(* IEC 61131-3 sources: veristc/veri-stc/tests/compiler-tests/positive, 6 files *)

(* ---- algo_blocks_fb.st ---- *)
(* ================================================================
   algo_blocks_fb.st
   原生 FUNCTION_BLOCK 版算法块库 + "不同变量调用相同算法功能" e2e

   与 FUNCTION 版（algo_blocks_lib.st / algo_blocks_multi_instance.st）
   同激励、同黄金时间线，可交叉验证两种实现一致。

   演示 FB 全部可用特性（P1 + v1.5）：
     - VAR_INPUT / VAR_OUTPUT（多输出：Q 与 QN、U 与 UI 与 ALM）
     - VAR 实例内持久状态（UI / E_OLD，FB_DATA 跨周期不清零）
     - VAR_IN_OUT 逐引用别名（TRACE：诊断量直写调用方全局）
     - 实例声明分离：rs1/rs2 同一份代码、独立数据段
     - IF/ELSIF/ELSE 控制流、表达式实参、命名实参（:=）
   限制：FB 体内不得声明成员实例（嵌套 FB 不支持，P1 范围外）。
   调用点在外部以 IEC 点号访问 inst.FIELD 读取字段（v1.5.1；编译器内部
   融合为不可书写的派生名 inst#FIELD，外部只能读 VAR_OUTPUT）。

   黄金时间线（数值列与 FUNCTION 版一致，t: rs1 rs2 sr1 sr2 | u1 ui1 |
   u2 ui2 | f1 f2，u 与 tr 恒等因 TRACE 别名）。列标签自 v1.5.1 起写作
   点号形式（rs1.Q / pid1.U / pid1.UI / fby1.Y …）指认"这一列来自哪个
   实例的哪个字段"；golden 文件随之只改标签文本，12 行数值逐列不变：
     t1 : 1 0 0 0 | 170 118 | 140 65  |  20   0
     t2 : 1 0 0 0 | 170 200 | 140 90  |  40   0
     t3 : 1 1 0 0 | 170 200 | 140 90  |  60   0
     t4 : 1 0 0 0 | 170 200 | 140 90  |  80   0
     t5 : 0 0 0 0 | 170 200 | 140 90  | 100  50
     t6 : 0 0 0 1 | 170 200 | 140 90  | 120 100
     t7 : 0 0 0 1 | 170 200 | 140 90  | 140 120
     t8 : 0 0 0 1 | 170 200 | 140 90  | 160 120
     t9 : 0 0 0 0 | 170 200 | 135 90  | 180 120
     t10: 0 0 0 0 | 170 200 | 125 90  | 200 120
     t11: 0 0 0 0 | 170 198 | 115 90  | 220 120
     t12: 0 0 0 0 | 158 184 | 105 90  | 240 120
   ================================================================ *)

(* ---- 实例声明：必须先于 POU 列表；每实例独立 FB_DATA ---- *)
VAR_GLOBAL
  rs1  : RS_FB;
  rs2  : RS_FB;
  sr1  : SR_FB;
  sr2  : SR_FB;
  pid1 : PID_FB;
  pid2 : PID_FB;
  fby1 : FBY_FB;
  fby2 : FBY_FB;
  trace1 : DINT;   (* pid1 的 VAR_IN_OUT 别名目标 *)
  trace2 : DINT;   (* pid2 的 VAR_IN_OUT 别名目标 *)
END_VAR

(* ---- RS：置位优先双稳态；Q 为实例持久状态 ---- *)
FUNCTION_BLOCK RS_FB
VAR_INPUT
  S : BOOL;
  R : BOOL;
END_VAR
VAR_OUTPUT
  Q  : BOOL;
  QN : BOOL;
END_VAR
  Q := S OR (Q AND NOT R);
  QN := NOT Q;
END_FUNCTION_BLOCK

(* ---- SR：复位优先双稳态 ---- *)
FUNCTION_BLOCK SR_FB
VAR_INPUT
  S : BOOL;
  R : BOOL;
END_VAR
VAR_OUTPUT
  Q  : BOOL;
  QN : BOOL;
END_VAR
  Q := (S OR Q) AND NOT R;
  QN := NOT Q;
END_FUNCTION_BLOCK

(* ---- PID：定点 PID，实例内持久 UI/E_OLD，KI 固定为 1；
       TRACE 为 VAR_IN_OUT 诊断别名，输出 U 同步写入调用方全局 ---- *)
FUNCTION_BLOCK PID_FB
VAR_INPUT
  E     : DINT;
  KP    : DINT;
  KD    : DINT;
  UI_LO : DINT;
  UI_HI : DINT;
  LO    : DINT;
  HI    : DINT;
END_VAR
VAR_OUTPUT
  U   : DINT;
  UI  : DINT;
  ALM : BOOL;
END_VAR
VAR_IN_OUT
  TRACE : DINT;
END_VAR
VAR
  DE    : DINT;
  V     : DINT;
  E_OLD : DINT;
END_VAR
  DE := E - E_OLD;
  V := UI + E;
  IF V > UI_HI THEN
    V := UI_HI;
  ELSIF V < UI_LO THEN
    V := UI_LO;
  END_IF;
  UI := V;
  U := KP * E + UI + KD * DE;
  IF U > HI THEN
    U := HI;
  ELSIF U < LO THEN
    U := LO;
  END_IF;
  IF U >= HI THEN
    ALM := TRUE;
  ELSE
    ALM := FALSE;
  END_IF;
  TRACE := U;
  E_OLD := E;
END_FUNCTION_BLOCK

(* ---- FBY：速率限制跟随；Y 为实例持久输出 ---- *)
FUNCTION_BLOCK FBY_FB
VAR_INPUT
  IN : DINT;
  DR : DINT;
END_VAR
VAR_OUTPUT
  Y : DINT;
END_VAR
VAR
  V : DINT;
END_VAR
  V := IN;
  IF V > Y + DR THEN
    V := Y + DR;
  ELSIF V < Y - DR THEN
    V := Y - DR;
  END_IF;
  Y := V;
END_FUNCTION_BLOCK

PROGRAM MAIN
VAR
  tick : DINT;
  in2  : DINT;
END_VAR
  tick := CycleCounter();

  (* 与 FUNCTION 版完全相同的激励时序 *)
  rs1(S := (tick = 1), R := (tick = 5));
  rs2(S := (tick = 3), R := (tick = 4));

  sr1(S := (tick = 2), R := (tick = 2));
  sr2(S := (tick = 6), R := (tick = 9));

  (* 同一份 PID 代码，两套增益/限值、两套独立状态与别名目标 *)
  pid1(E := 130 - tick * 12, KP := 1, KD := 1,
       UI_LO := 0, UI_HI := 200, LO := 0, HI := 170,
       TRACE := trace1);
  pid2(E := 70 - tick * 5, KP := 2, KD := 1,
       UI_LO := 0, UI_HI := 90, LO := 0, HI := 140,
       TRACE := trace2);

  fby1(IN := tick * 30, DR := 20);
  IF tick > 4 THEN
    in2 := 120;
  ELSE
    in2 := 0;
  END_IF;
  fby2(IN := in2, DR := 50);

  PRINT('FB t=', tick, ' rs1.Q,=', rs1.Q, ' rs2.Q,=', rs2.Q,
        ' sr1.Q,=', sr1.Q, ' sr2.Q,=', sr2.Q,
        ' pid1.U,=', pid1.U, ' pid1.UI,=', pid1.UI,
        ' pid2.U,=', pid2.U, ' pid2.UI,=', pid2.UI,
        ' fby1.Y,=', fby1.Y, ' fby2.Y,=', fby2.Y,
        ' trace1,=', trace1, ' trace2,=', trace2, '\n');
END_PROGRAM

(* ---- in_out_alias_field.st ---- *)
(* ================================================================
   positive/in_out_alias_field.st  --  别名目标可以是实例数据字段

   a2.ACC 绑定到 a1.LAST（expand_instances 展开出的扁平全局字段），
   即"跨实例逐引用"：a2 的写直接落在 a1 的输出字段存储上，
   与 a1 自己的读写共享同一地址。合法 ⇒ 编译器必须接受。
   ================================================================ *)

VAR_GLOBAL
  t : DINT;
  tick : DINT;
  a1 : FB_INC;
  a2 : FB_INC;
END_VAR

FUNCTION_BLOCK FB_INC
VAR_INPUT
  K : DINT;
END_VAR
VAR_OUTPUT
  LAST : DINT;
END_VAR
VAR_IN_OUT
  ACC : DINT;
END_VAR
  LAST := ACC;
  ACC := ACC + K;
END_FUNCTION_BLOCK

PROGRAM MAIN
  tick := CycleCounter();
  t := tick;
  a1(ACC := t, K := 1);
  a2(ACC := a1.LAST, K := 5);
  PRINT('t', t, a1.LAST, a2.LAST);
END_PROGRAM

(* ---- algo_blocks_multi_instance.st ---- *)
(* ================================================================
   algo_blocks_multi_instance.st
   测试用例：不同的变量调用相同的算法功能（多实例复用）

   内联库：tests/st-examples/algo_blocks_lib.st
   （VeriSTC 无库链接机制，库文本由上游预处理器内联，此处手工内联）

   每个算法块均有 2 个实例，实例之间变量完全独立：
     RS(q1)/RS(q2)   SR(q1)/SR(q2)
     PID(e1,ui1,de1,u1) / PID(e2,ui2,de2,u2)
     FBY(in->f1) / FBY(in->f2)
   跨周期状态全部放 VAR_GLOBAL 并由调用方写回。

   12 周期金标准（t: rs1 rs2 sr1 sr2 | u1 ui1 | u2 ui2 | f1 f2）
     t1 : 1 0 0 0 | 170 118 | 140 65  |  20   0
     t2 : 1 0 0 0 | 170 200 | 140 90  |  40   0
     t3 : 1 1 0 0 | 170 200 | 140 90  |  60   0
     t4 : 1 0 0 0 | 170 200 | 140 90  |  80   0
     t5 : 0 0 0 0 | 170 200 | 140 90  | 100  50
     t6 : 0 0 0 1 | 170 200 | 140 90  | 120 100
     t7 : 0 0 0 1 | 170 200 | 140 90  | 140 120
     t8 : 0 0 0 1 | 170 200 | 140 90  | 160 120
     t9 : 0 0 0 0 | 170 200 | 135 90  | 180 120
     t10: 0 0 0 0 | 170 200 | 125 90  | 200 120
     t11: 0 0 0 0 | 170 198 | 115 90  | 220 120
     t12: 0 0 0 0 | 158 184 | 105 90  | 240 120
   ================================================================ *)

VAR_GLOBAL
  rs1_q  : BOOL;
  rs2_q  : BOOL;
  sr1_q  : BOOL;
  sr2_q  : BOOL;
  pid1_ui   : DINT;
  pid1_eold : DINT;
  pid2_ui   : DINT;
  pid2_eold : DINT;
  fby1_out : DINT;
  fby2_out : DINT;
END_VAR

(* ---------------- 库：algo_blocks_lib.st 内联开始 ---------------- *)

FUNCTION RS : BOOL
VAR_INPUT
  Q_old : BOOL;
  S : BOOL;
  R : BOOL;
END_VAR
  RS := S OR (Q_old AND NOT R);
END_FUNCTION

FUNCTION SR : BOOL
VAR_INPUT
  Q_old : BOOL;
  S : BOOL;
  R : BOOL;
END_VAR
  SR := (S OR Q_old) AND NOT R;
END_FUNCTION

FUNCTION PID_UI : DINT
VAR_INPUT
  E  : DINT;
  UI : DINT;
  KI : DINT;
  LO : DINT;
  HI : DINT;
END_VAR
VAR
  V : DINT;
END_VAR
  V := UI + KI * E;
  IF V > HI THEN
    V := HI;
  ELSIF V < LO THEN
    V := LO;
  END_IF;
  PID_UI := V;
END_FUNCTION

FUNCTION PID_OUT : DINT
VAR_INPUT
  E   : DINT;
  UI  : DINT;
  DE  : DINT;
  KP  : DINT;
  KD  : DINT;
  LO  : DINT;
  HI  : DINT;
END_VAR
VAR
  U : DINT;
END_VAR
  U := KP * E + UI + KD * DE;
  IF U > HI THEN
    U := HI;
  ELSIF U < LO THEN
    U := LO;
  END_IF;
  PID_OUT := U;
END_FUNCTION

FUNCTION FBY : DINT
VAR_INPUT
  IN  : DINT;
  PRE : DINT;
  DR  : DINT;
END_VAR
VAR
  Q : DINT;
END_VAR
  Q := IN;
  IF Q > PRE + DR THEN
    Q := PRE + DR;
  ELSIF Q < PRE - DR THEN
    Q := PRE - DR;
  END_IF;
  FBY := Q;
END_FUNCTION

(* ---------------- 库内联结束 ---------------- *)

PROGRAM MAIN
VAR
  tick  : DINT;
  rs1_s : BOOL;
  rs1_r : BOOL;
  rs2_s : BOOL;
  rs2_r : BOOL;
  sr1_s : BOOL;
  sr1_r : BOOL;
  sr2_s : BOOL;
  sr2_r : BOOL;
  e1  : DINT;
  de1 : DINT;
  u1  : DINT;
  e2  : DINT;
  de2 : DINT;
  u2  : DINT;
  in1 : DINT;
  in2 : DINT;
  fby1_q : DINT;
  fby2_q : DINT;
END_VAR
  tick := CycleCounter();

  (* ---- 激励 ---- *)
  rs1_s := tick = 1;
  rs1_r := tick = 5;
  rs2_s := tick = 3;
  rs2_r := tick = 4;
  sr1_s := tick = 2;
  sr1_r := tick = 2;
  sr2_s := tick = 6;
  sr2_r := tick = 9;

  (* ---- RS：同一功能，两套变量 ---- *)
  rs1_q := RS(rs1_q, rs1_s, rs1_r);
  rs2_q := RS(rs2_q, rs2_s, rs2_r);

  (* ---- SR：同一功能，另两套变量 ---- *)
  sr1_q := SR(sr1_q, sr1_s, sr1_r);
  sr2_q := SR(sr2_q, sr2_s, sr2_r);

  (* ---- PID 实例 1：e1 = 130 - 12t, Kp=Ki=Kd=1, UI限[0,200], U限[0,170] ---- *)
  e1  := 130 - tick * 12;
  de1 := e1 - pid1_eold;
  pid1_ui := PID_UI(e1, pid1_ui, 1, 0, 200);
  u1  := PID_OUT(e1, pid1_ui, de1, 1, 1, 0, 170);
  pid1_eold := e1;

  (* ---- PID 实例 2：e2 = 70 - 5t, Kp=2,Kd=1, UI限[0,90], U限[0,140] ---- *)
  e2  := 70 - tick * 5;
  de2 := e2 - pid2_eold;
  pid2_ui := PID_UI(e2, pid2_ui, 1, 0, 90);
  u2  := PID_OUT(e2, pid2_ui, de2, 2, 1, 0, 140);
  pid2_eold := e2;

  (* ---- FBY 实例 1：in1 = 30t 斜坡, 速率限 20 ---- *)
  in1 := tick * 30;
  fby1_q := FBY(in1, fby1_out, 20);
  fby1_out := fby1_q;

  (* ---- FBY 实例 2：t<=4 时 in2=0，之后跳变 120, 速率限 50 ---- *)
  IF tick > 4 THEN
    in2 := 120;
  ELSE
    in2 := 0;
  END_IF;
  fby2_q := FBY(in2, fby2_out, 50);
  fby2_out := fby2_q;

  PRINT('ALG t=', tick, ' rs1=', rs1_q, ' rs2=', rs2_q,
        ' sr1=', sr1_q, ' sr2=', sr2_q,
        ' u1=', u1, ' ui1=', pid1_ui,
        ' u2=', u2, ' ui2=', pid2_ui,
        ' f1=', fby1_out, ' f2=', fby2_out, '\n');
END_PROGRAM

(* ---- function_basic.st ---- *)
(* Positive test: valid FUNCTION with local variable and IF control flow. *)

FUNCTION AddOne : DINT
VAR_INPUT
  val : DINT;
END_VAR
VAR
  r : DINT;
END_VAR
  IF val > 0 THEN
    r := val + 1;
  ELSE
    r := 0;
  END_IF;
  AddOne := r;
END_FUNCTION

PROGRAM function_basic
VAR
  result : DINT;
END_VAR
  result := AddOne(41);
  PRINT('result=', result, '\n');
END_PROGRAM

(* ---- minimal_assign.st ---- *)
(* Positive test: minimal valid program. *)

PROGRAM minimal_assign
VAR
  x : DINT;
END_VAR
  x := 42;
  PRINT('x=', x, '\n');
END_PROGRAM

(* ---- real_literals.st ---- *)
(* Positive test: REAL decimal literals.

   Each literal is stored straight into its own REAL local, so the code
   section holds one F32_CONST + LOCAL_SET pair per row and nothing else.
   The expected single-precision bit patterns are checked byte by byte by
   step 3 of run_compiler_tests.sh (f32 immediates on the wire). *)

PROGRAM real_literals
VAR
  v00 : REAL;
  v01 : REAL;
  v02 : REAL;
  v03 : REAL;
  v04 : REAL;
  v05 : REAL;
  v06 : REAL;
  v07 : REAL;
  v08 : REAL;
  v09 : REAL;
  v10 : REAL;
  v11 : REAL;
  v12 : REAL;
  v13 : REAL;
END_VAR
  v00 := 1.5;
  v01 := 0.1;
  v02 := -0.1;
  v03 := 3.14159265;
  v04 := 16777217.0;
  v05 := 0.33333333333333;
  v06 := 1.0e6;
  v07 := 2.5e-1;
  v08 := -1.5;
  v09 := 0.0000001;
  v10 := 1.0e-9;
  v11 := 100.0;
  v12 := 0.0;
  v13 := -273.15;
END_PROGRAM
